// LS Electric XG5000 project: PLC_PC_Test
// PLC LSPLC
// module base 0 slot 0: 입출력 모듈:XBM-DN32H (DC 24V입력/TR 출력, 32점)
// module base 0 slot 2: 위치결정 모듈:XBF-PD02A (위치결정 펄스(LD)출력형, 2축)

PROGRAM PcControll (task: 스캔 프로그램)

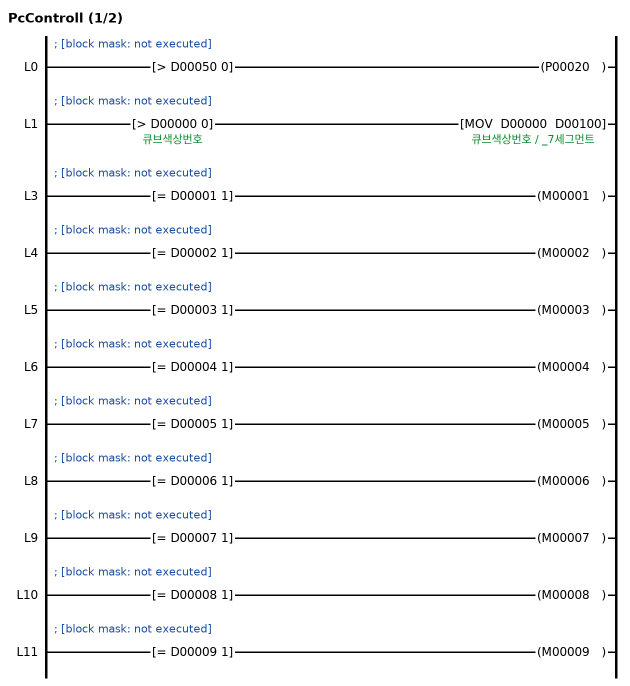
; L0 (block mask: not executed)
LOAD>     D00050 0
OUT       P00020
; L1 (block mask: not executed)
LOAD>     D00000 0	// 큐브색상번호
MOV       D00000 D00100	// 큐브색상번호 / _7세그먼트
; L3 (block mask: not executed)
LOAD=     D00001 1
OUT       M00001
; L4 (block mask: not executed)
LOAD=     D00002 1
OUT       M00002
; L5 (block mask: not executed)
LOAD=     D00003 1
OUT       M00003
; L6 (block mask: not executed)
LOAD=     D00004 1
OUT       M00004
; L7 (block mask: not executed)
LOAD=     D00005 1
OUT       M00005
; L8 (block mask: not executed)
LOAD=     D00006 1
OUT       M00006
; L9 (block mask: not executed)
LOAD=     D00007 1
OUT       M00007
; L10 (block mask: not executed)
LOAD=     D00008 1
OUT       M00008
; L11 (block mask: not executed)
LOAD=     D00009 1
OUT       M00009

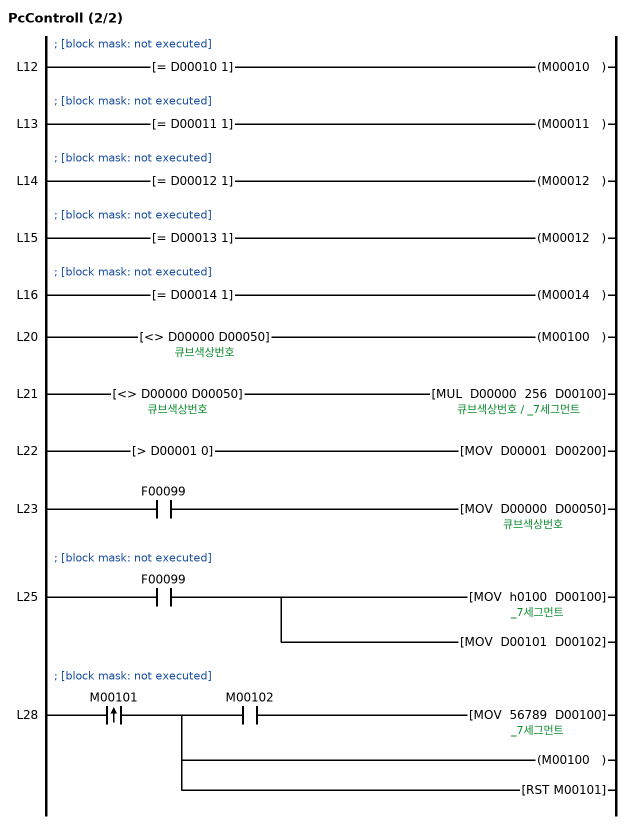
; L12 (block mask: not executed)
LOAD=     D00010 1
OUT       M00010
; L13 (block mask: not executed)
LOAD=     D00011 1
OUT       M00011
; L14 (block mask: not executed)
LOAD=     D00012 1
OUT       M00012
; L15 (block mask: not executed)
LOAD=     D00013 1
OUT       M00012
; L16 (block mask: not executed)
LOAD=     D00014 1
OUT       M00014
; L20
LOAD<>    D00000 D00050	// 큐브색상번호
OUT       M00100
; L21
LOAD<>    D00000 D00050	// 큐브색상번호
MUL       D00000 256 D00100	// 큐브색상번호 / _7세그먼트
; L22
LOAD>     D00001 0
MOV       D00001 D00200
; L23
LOAD      F00099
MOV       D00000 D00050	// 큐브색상번호
; L25 (block mask: not executed)
LOAD      F00099
MOV       h0100 D00100	// _7세그먼트
MOV       D00101 D00102
; L28 (block mask: not executed)
LOADP     M00101
MPUSH
AND       M00102
MOV       56789 D00100	// _7세그먼트
MPOP
OUT       M00100
RST       M00101